(*
SPDX-FileCopyrightText: c 2026 Oleksandr Tiutyk <trofimich@gmail.com>
SPDX-License-Identifier: MIT
License: https://opensource.org/license/mit
*)

(*!
<summary>Checks absolute dispersion and independent output clamps.</summary>
<description>
Owns a generator used by one PLC task. Each run checks the same bounds against fresh samples.
The runner binds assertions to the instance address. Keep the instance at that address for its run.
</description>
*)

{attribute 'no_assign'}
{attribute 'no_explicit_call' := 'do not call this function block directly'}
FUNCTION_BLOCK RandomAbsoluteDispersionTest EXTENDS TOF_Testing.SingleCycleTest
VAR_STAT
	{attribute 'hide'}
	_ClassName : STRING := __POUNAME();
END_VAR
VAR
	_Random : TOF_Core.Random;
END_VAR

//! <summary>Checks zero dispersion and bounds that must clamp independently of the generated sample.</summary>
METHOD PROTECTED ExecuteTest
VAR
	value : LREAL;
	i : INT;
END_VAR
value := _Random.GetWithDispersion(baseValue := LREAL#12.5, dispersion := LREAL#0.0);
Assert.ThatLongReal(actual := value, message := "Zero dispersion must return the base").ToBe(expected := LREAL#12.5);

value := _Random.GetWithDispersion(baseValue := LREAL#100.0, dispersion := LREAL#10.0, minValue := LREAL#120.0);
Assert.ThatLongReal(
	actual := value,
	message := "Lower bound alone must clamp any sample"
).ToBe(expected := LREAL#120.0);

value := _Random.GetWithDispersion(baseValue := LREAL#100.0, dispersion := LREAL#10.0, maxValue := LREAL#80.0);
Assert.ThatLongReal(actual := value, message := "Upper bound alone must clamp any sample").ToBe(expected := LREAL#80.0);

FOR i := 1 TO 21 DO
	value := _Random.GetWithDispersion(baseValue := LREAL#100.0, dispersion := LREAL#10.0);
	Assert.ThatLongReal(
	actual := value,
	message := "Absolute dispersion sample below 90"
).IsGreaterThanOrEquals(
		expected := LREAL#90.0
	);
	Assert.ThatLongReal(
	actual := value,
	message := "Absolute dispersion sample above 110"
).IsLessThanOrEquals(
		expected := LREAL#110.0
	);
END_FOR
END_METHOD

//! <summary>Borrows the concrete class name. Callers must not modify it.</summary>
{attribute 'monitoring' := 'call'}
PROPERTY ClassName : REFERENCE TO STRING
GET
ClassName REF= _ClassName;
END_GET
END_PROPERTY

//! <summary>Borrows the compiler-initialized namespace name. Callers must not modify it.</summary>
{attribute 'monitoring' := 'call'}
PROPERTY NamespaceName : REFERENCE TO STRING
GET
NamespaceName REF= CurrentNamespace.Name;
END_GET
END_PROPERTY

//! <summary>Reports the concrete instance size in bytes.</summary>
{attribute 'monitoring' := 'call'}
PROPERTY SelfSize : ULINT
GET
SelfSize := XSIZEOF(THIS^);
END_GET
END_PROPERTY

END_FUNCTION_BLOCK

(* stored: Version 1.1.0.1
   POU RandomAbsoluteDispersionTest: Id {70f7b36d-6374-4f42-9bd6-22c0fd1f07a5}, SpecialFunc None
   Method ExecuteTest: Id {bd814188-2ec2-4d28-93fa-70a22c7528d5}
   Property ClassName: Id {5e788ffb-fa0c-4d12-80a1-75242a6282ab}
   Get Get: Id {1802a401-5f28-452b-8eef-a98603de327c}
   Property NamespaceName: Id {fdf9a300-b1e4-42ab-9200-35ae2b508d3b}
   Get Get: Id {bb691c65-f18e-4349-b32e-39d62d4f0b0e}
   Property SelfSize: Id {7ce4fc59-3452-417e-a4cb-a42aef41defb}
   Get Get: Id {31dc69fe-f1ee-4efb-95c9-aa6366cbc377} *)
